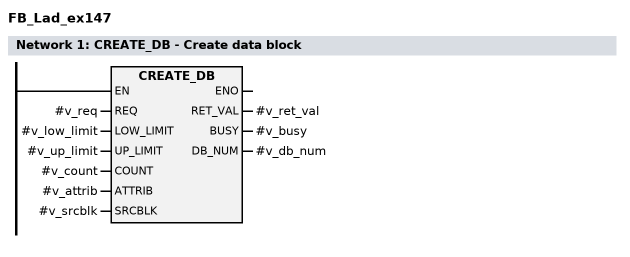
   #v_ret_val := CREATE_DB(REQ := #v_req,
                           LOW_LIMIT := #v_low_limit,
                           UP_LIMIT := #v_up_limit,
                           COUNT := #v_count,
                           ATTRIB := #v_attrib,
                           SRCBLK := #v_srcblk,
                           BUSY => #v_busy,
                           DB_NUM => #v_db_num);
END_REGION
END_FUNCTION_BLOCK

FUNCTION_BLOCK "FB_Lad_ex150"   // FB54, LAD
{ S7_Optimized_Access := 'TRUE' }
   VAR_INPUT
      v_req : Bool;
      v_db_number : DB_ANY;
   END_VAR
   VAR_OUTPUT
      v_ret_val : Int;
      v_db_length : UDInt;
      v_attrib : Byte;
   END_VAR
BEGIN

REGION Network 1: ATTR_DB - Read data block attribute
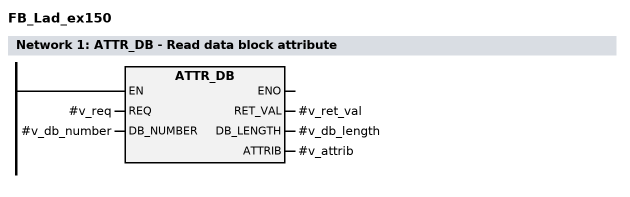
   #v_ret_val := ATTR_DB(REQ := #v_req,
                         DB_NUMBER := #v_db_number,
                         DB_LENGTH => #v_db_length,
                         ATTRIB => #v_attrib);
END_REGION
END_FUNCTION_BLOCK

FUNCTION_BLOCK "FB_Lad_ex151"   // FB55, LAD
{ S7_Optimized_Access := 'TRUE' }
   VAR_INPUT
      v_req : Bool;
      v_db_number : UInt;
   END_VAR
   VAR_OUTPUT
      v_ret_val : Int;
      v_busy : Bool;
   END_VAR
BEGIN

REGION Network 1: DELETE_DB - Delete data block
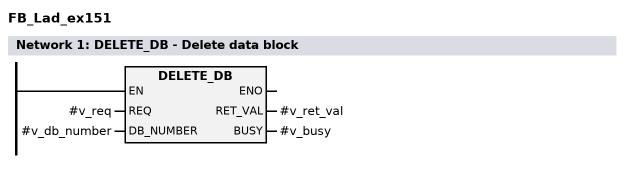
   #v_ret_val := DELETE_DB(REQ := #v_req, DB_NUMBER := #v_db_number, BUSY => #v_busy);
END_REGION
END_FUNCTION_BLOCK

FUNCTION_BLOCK "FB_Lad_ex154"   // FB56, LAD
{ S7_Optimized_Access := 'TRUE' }
   VAR_INPUT
      v_ioid : Byte;
      v_addr : Word;
      v_ret_val : Int;
   END_VAR
   VAR_OUTPUT
      v_hwid : Hw_Io;
   END_VAR
BEGIN

REGION Network 1: LOG2MOD - Determine the hardware identifier from addressing of STEP 7 V5.5 SPx
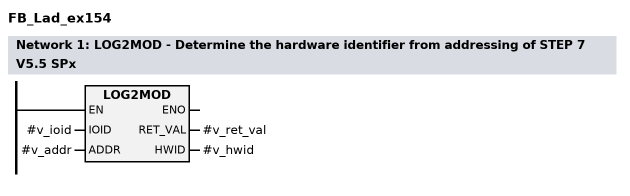
   #v_ret_val := LOG2MOD(IOID := #v_ioid, ADDR := #v_addr, HWID => #v_hwid);
END_REGION
END_FUNCTION_BLOCK

FUNCTION_BLOCK "FB_Lad_ex155"   // FB57, LAD
{ S7_Optimized_Access := 'TRUE' }
   VAR_INPUT
      v_addr : Variant;
      v_ret_val : Int;
   END_VAR
   VAR_OUTPUT
      v_laddr : Hw_Io;
   END_VAR
BEGIN

REGION Network 1: IO2MOD - Determine hardware identifier from an IO address
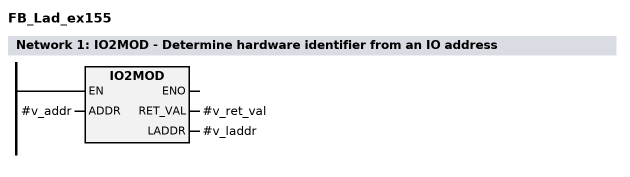
   #v_ret_val := IO2MOD(ADDR := #v_addr, LADDR => #v_laddr);
END_REGION
END_FUNCTION_BLOCK

FUNCTION_BLOCK "FB_Lad_ex156"   // FB58, LAD
{ S7_Optimized_Access := 'TRUE' }
   VAR_INPUT
      v_laddr : Hw_Io;
      v_ret_val : Int;
   END_VAR
   VAR_OUTPUT
      v_piaddr : UDInt;
      v_picount : UInt;
      v_pqaddr : UDInt;
      v_pqcount : UInt;
   END_VAR
BEGIN

REGION Network 1: RD_ADDR - Determine IO addresses from the hardware identifier
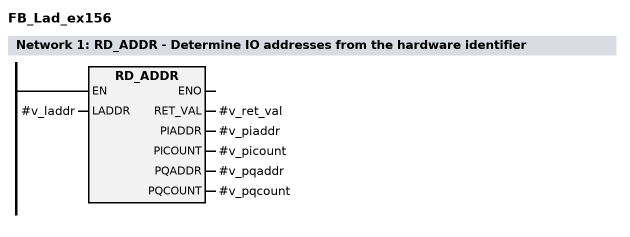
   #v_ret_val := RD_ADDR(LADDR := #v_laddr,
                         PIADDR => #v_piaddr,
                         PICount => #v_picount,
                         PQADDR => #v_pqaddr,
                         PQCount => #v_pqcount);
END_REGION
END_FUNCTION_BLOCK

FUNCTION_BLOCK "FB_Lad_ex157"   // FB59, LAD
{ S7_Optimized_Access := 'TRUE' }
   VAR_INPUT
      v_master : Int;
      v_station : Int;
      v_slot : Int;
      v_subslot : Int;
      v_ret_val : Int;
   END_VAR
   VAR_OUTPUT
      v_laddr : Hw_Io;
   END_VAR
BEGIN

REGION Network 1: GEO_LOG - Determine hardware identifier from slot
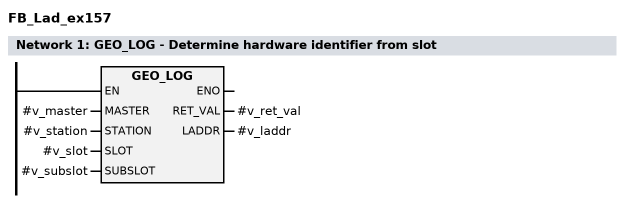
   #v_ret_val := GEO_LOG(MASTER := #v_master,
                         STATION := #v_station,
                         SLOT := #v_slot,
                         SUBSLOT := #v_subslot,
                         LADDR => #v_laddr);
END_REGION
END_FUNCTION_BLOCK

FUNCTION_BLOCK "FB_Lad_ex158"   // FB60, LAD
{ S7_Optimized_Access := 'TRUE' }
   VAR_INPUT
      v_laddr : Hw_Io;
      v_ret_val : Int;
   END_VAR
   VAR_OUTPUT
      v_area : Int;
      v_master : Int;
      v_station : Int;
      v_slot : Int;
      v_subslot : Int;
      v_offset : Int;
   END_VAR
BEGIN

REGION Network 1: LOG_GEO - Determine slot from hardware identifier
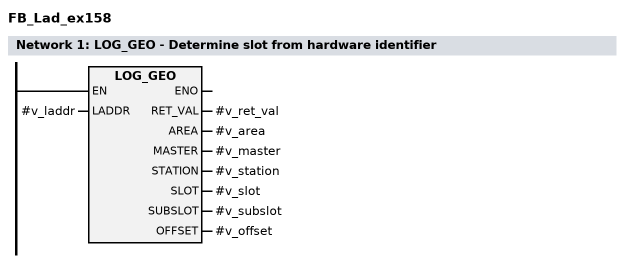
   #v_ret_val := LOG_GEO(LADDR := #v_laddr,
                         AREA => #v_area,
                         MASTER => #v_master,
                         STATION => #v_station,
                         SLOT => #v_slot,
                         SUBSLOT => #v_subslot,
                         OFFSET => #v_offset);
END_REGION
END_FUNCTION_BLOCK

FUNCTION_BLOCK "FB_Lad_ex160"   // FB61, LAD
{ S7_Optimized_Access := 'TRUE' }
   VAR_INPUT
      v_subnetid : Byte;
      v_rack : Word;
      v_slot : Word;
      v_subslot : Byte;
      v_subaddr : Word;
      v_ret_val : Int;
   END_VAR
   VAR_OUTPUT
      v_ioid : Byte;
      v_laddr : Hw_Module;
   END_VAR
BEGIN

REGION Network 1: GADR_LGC - Determine hardware identifier from slot and offset in the user data address area
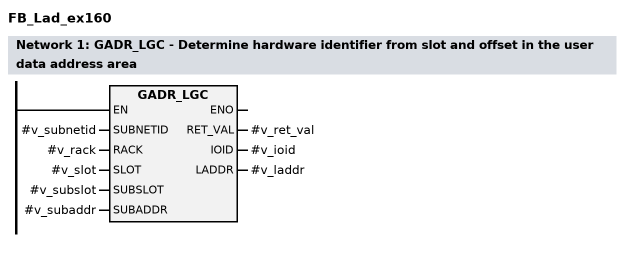
   #v_ret_val := GADR_LGC(SUBNETID := #v_subnetid,
                          RACK := #v_rack,
                          SLOT := #v_slot,
                          SUBSLOT := #v_subslot,
                          SUBADDR := #v_subaddr,
                          IOID => #v_ioid,
                          LADDR => #v_laddr);
END_REGION
END_FUNCTION_BLOCK

FUNCTION_BLOCK "FB_Lad_ex161"   // FB62, LAD
{ S7_Optimized_Access := 'TRUE' }
   VAR_INPUT
      v_ioid : Byte;
      v_laddr : Hw_Module;
      v_ret_val : Int;
   END_VAR
   VAR_OUTPUT
      v_area : Byte;
      v_rack : Word;
      v_slot : Word;
      v_subaddr : Word;
   END_VAR
BEGIN

REGION Network 1: LGC_GADR - Determine slot from hardware identifier
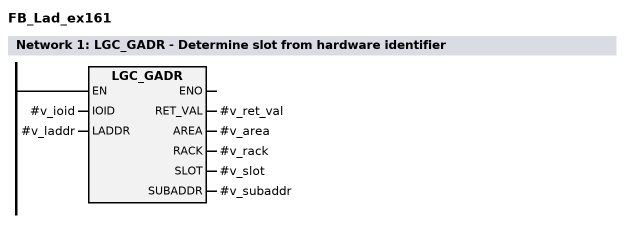
   #v_ret_val := LGC_GADR(IOID := #v_ioid,
                          LADDR := #v_laddr,
                          AREA => #v_area,
                          RACK => #v_rack,
                          SLOT => #v_slot,
                          SUBADDR => #v_subaddr);
END_REGION
END_FUNCTION_BLOCK

FUNCTION_BLOCK "FB_Lad_ws001"   // FB63, LAD
{ S7_Optimized_Access := 'TRUE' }
   VAR_INPUT
      v_ctrl_db : DB_WWW;
   END_VAR
   VAR_OUTPUT
      v_ret_val : Int;
   END_VAR
BEGIN

REGION Network 1: WWW - Synchronizing user pages
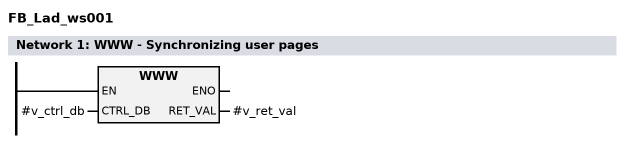
   #v_ret_val := WWW(CTRL_DB := #v_ctrl_db);
END_REGION
END_FUNCTION_BLOCK

FUNCTION_BLOCK "FB_Lad_ex025"   // FB64, LAD
{ S7_Optimized_Access := 'TRUE' }
   VAR_INPUT
      v_n : Int;
      v_ret_val : Word;
   END_VAR
   VAR_IN_OUT
      v_in : Variant;
      v_out : Variant;
   END_VAR
BEGIN

REGION Network 1: ATH - Convert ASCII string to hexadecimal number
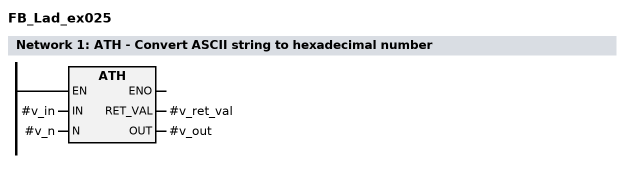
   #v_ret_val := ATH(IN := #v_in, N := #v_n, OUT => #v_out);
END_REGION
END_FUNCTION_BLOCK

FUNCTION_BLOCK "FB_Lad_ex026"   // FB65, LAD
{ S7_Optimized_Access := 'TRUE' }
   VAR_INPUT
      v_n : UInt;
      v_ret_val : Word;
   END_VAR
   VAR_IN_OUT
      v_in : Variant;
      v_out : Variant;
   END_VAR
BEGIN

REGION Network 1: HTA - Convert hexadecimal number to ASCII string
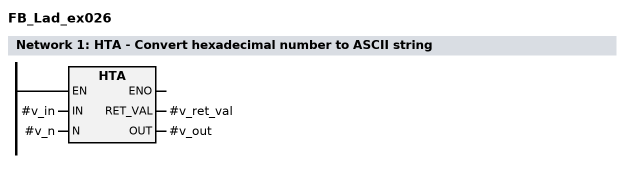
   #v_ret_val := HTA(IN := #v_in, N := #v_n, OUT => #v_out);
END_REGION
END_FUNCTION_BLOCK

FUNCTION_BLOCK "FB_Lad_ex036"   // FB66, LAD
{ S7_Optimized_Access := 'TRUE' }
   VAR_INPUT
      v_size : DInt;
      v_out : WString;
   END_VAR
   VAR_IN_OUT
      v_variable : Array[0..99] of Byte;
   END_VAR
BEGIN

REGION Network 1: GetSymbolName - Read out a tag on the input parameter
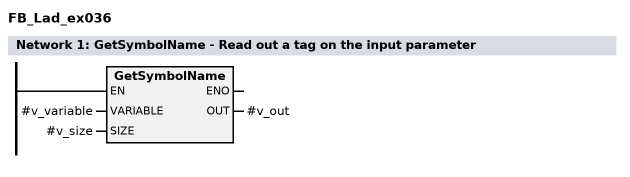
   // no SCL statement known for GetSymbolName: written as a call
   #v_out := GetSymbolName(variable := #v_variable, size := #v_size);
END_REGION
END_FUNCTION_BLOCK

FUNCTION_BLOCK "FB_Lad_ex060"   // FB67, LAD
{ S7_Optimized_Access := 'TRUE' }
   VAR_INPUT
      v_laddr : Hw_Io;
      v_ret_val : Int;
   END_VAR
   VAR_IN_OUT
      v_record : Variant;
   END_VAR
BEGIN

REGION Network 1: DPRD_DAT - Read consistent data of a DP standard slave
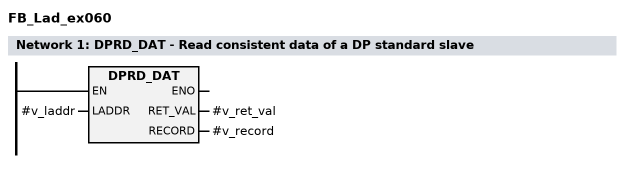
   #v_ret_val := DPRD_DAT(LADDR := #v_laddr, RECORD => #v_record);
END_REGION
END_FUNCTION_BLOCK

FUNCTION_BLOCK "FB_Lad_ex065"   // FB68, LAD
{ S7_Optimized_Access := 'TRUE' }
   VAR_INPUT
      v_req : Bool;
      v_laddr : Hw_DpSlave;
      v_ret_val : DInt;
   END_VAR
   VAR_OUTPUT
      v_busy : Bool;
   END_VAR
   VAR_IN_OUT
      v_record : Variant;
   END_VAR
BEGIN

REGION Network 1: DPNRM_DG - Read diagnostics data from a DP slave
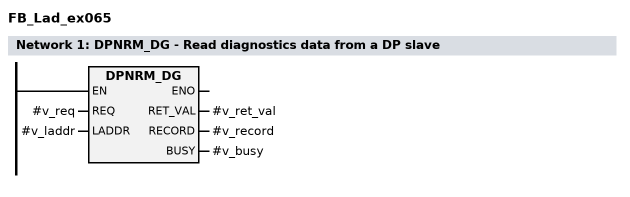
   #v_ret_val := DPNRM_DG(REQ := #v_req, LADDR := #v_laddr, RECORD => #v_record, BUSY => #v_busy);
END_REGION
END_FUNCTION_BLOCK

FUNCTION_BLOCK "FB_Lad_ex097"   // FB69, LAD
{ S7_Optimized_Access := 'TRUE' }
   VAR_INPUT
      v_req : Bool;
      v_laddr : Hw_Io;
      v_recnum : Byte;
      v_ret_val : Int;
   END_VAR
   VAR_OUTPUT
      v_busy : Bool;
   END_VAR
   VAR_IN_OUT
      v_record : Variant;
   END_VAR
BEGIN

REGION Network 1: RD_DPARA - Read module data record asynchronously
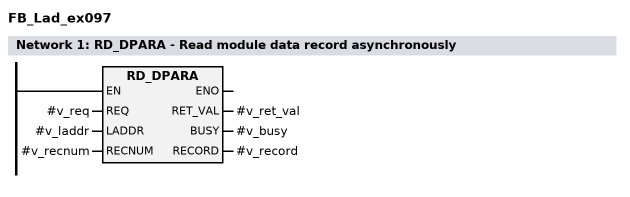
   #v_ret_val := RD_DPARA(REQ := #v_req,
                          LADDR := #v_laddr,
                          RECNUM := #v_recnum,
                          BUSY => #v_busy,
                          RECORD => #v_record);
END_REGION
END_FUNCTION_BLOCK

FUNCTION_BLOCK "FB_Lad_ex098"   // FB70, LAD
{ S7_Optimized_Access := 'TRUE' }
   VAR_INPUT
      v_ioid : Byte;
      v_laddr : Hw_Io;
      v_recnum : Byte;
      v_ret_val : Int;
   END_VAR
   VAR_IN_OUT
      v_record : Variant;
   END_VAR
BEGIN

REGION Network 1: RD_DPARM - Read data record from configured system data
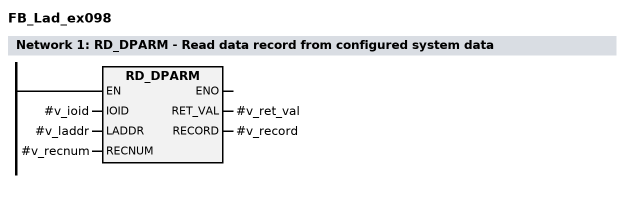
   #v_ret_val := RD_DPARM(IOID := #v_ioid, LADDR := #v_laddr, RECNUM := #v_recnum, RECORD => #v_record);
END_REGION
END_FUNCTION_BLOCK

FUNCTION_BLOCK "FB_Lad_ex124"   // FB71, LAD
{ S7_Optimized_Access := 'TRUE' }
   VAR_INPUT
      v_ret_val : Int;
   END_VAR
   VAR_IN_OUT
      v_top_si : Array[0..99] of Byte;
      v_start_up_si : Array[0..99] of Byte;
   END_VAR
BEGIN

REGION Network 1: RD_SINFO - Read current OB start information
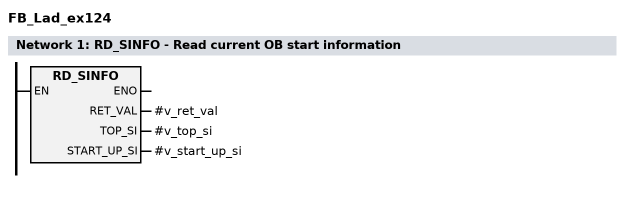
   #v_ret_val := RD_SINFO(TOP_SI => #v_top_si, START_UP_SI => #v_start_up_si);
END_REGION
END_FUNCTION_BLOCK

FUNCTION_BLOCK "FB_Lad_ex148"   // FB72, LAD
{ S7_Optimized_Access := 'TRUE' }
   VAR_INPUT
      v_req : Bool;
      v_ret_val : Int;
   END_VAR
   VAR_OUTPUT
      v_busy : Bool;
   END_VAR
   VAR_IN_OUT
      v_srcblk : Variant;
      v_dstblk : Variant;
   END_VAR
BEGIN

REGION Network 1: READ_DBL - Read from data block in the load memory
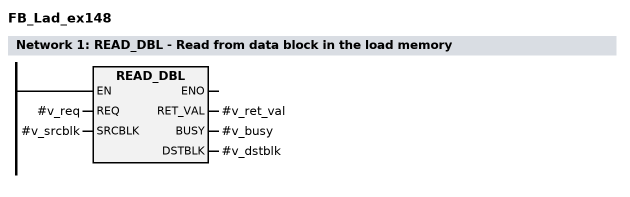
   #v_ret_val := READ_DBL(REQ := #v_req, SRCBLK := #v_srcblk, BUSY => #v_busy, DSTBLK => #v_dstblk);
END_REGION
END_FUNCTION_BLOCK

FUNCTION_BLOCK "FB_Lad_ex149"   // FB73, LAD
{ S7_Optimized_Access := 'TRUE' }
   VAR_INPUT
      v_req : Bool;
      v_ret_val : Int;
   END_VAR
   VAR_OUTPUT
      v_busy : Bool;
   END_VAR
   VAR_IN_OUT
      v_srcblk : Variant;
      v_dstblk : Variant;
   END_VAR
BEGIN

REGION Network 1: WRIT_DBL - Write to data block in the load memory
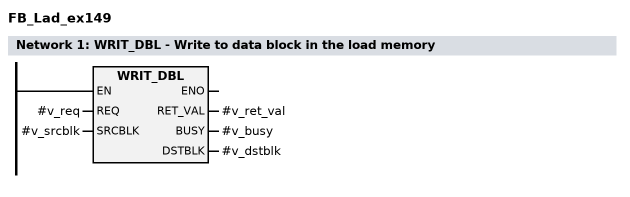
   #v_ret_val := WRIT_DBL(REQ := #v_req, SRCBLK := #v_srcblk, BUSY => #v_busy, DSTBLK => #v_dstblk);
END_REGION
END_FUNCTION_BLOCK

FUNCTION_BLOCK "FB_Lad_ou010"   // FB74, LAD
{ S7_Optimized_Access := 'TRUE' }
   VAR_INPUT
      v_req : Bool;
      v_id : Conn_Ouc;
   END_VAR
   VAR_OUTPUT
      v_done : Bool;
      v_busy : Bool;
      v_error : Bool;
      v_status : Word;
   END_VAR
   VAR_IN_OUT
      v_connect : TCON_Param;
   END_VAR
   VAR
      inst : TCON;
   END_VAR
BEGIN

REGION Network 1: TCON - Establish communication connection
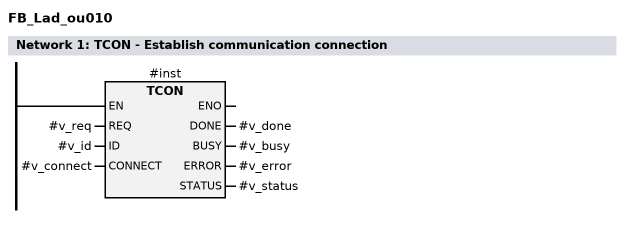
   #inst(REQ := #v_req,   // TCON
         ID := #v_id,
         CONNECT := #v_connect,
         DONE => #v_done,
         BUSY => #v_busy,
         ERROR => #v_error,
         STATUS => #v_status);
END_REGION
END_FUNCTION_BLOCK

FUNCTION_BLOCK "FB_Lad_ou002"   // FB75, LAD
{ S7_Optimized_Access := 'TRUE' }
   VAR_INPUT
      v_req : Bool;
      v_cont : Bool;
      v_len : UDInt;
   END_VAR
   VAR_OUTPUT
      v_done : Bool;
      v_busy : Bool;
      v_error : Bool;
      v_status : Word;
   END_VAR
   VAR_IN_OUT
      v_connect : Array[0..99] of Byte;
      v_data : Array[0..99] of Byte;
      v_addr : Array[0..99] of Byte;
      v_com_rst : Bool;
   END_VAR
   VAR
      inst : TSEND_C;
   END_VAR
BEGIN

REGION Network 1: TSEND_C - Establishing a connection and sending data
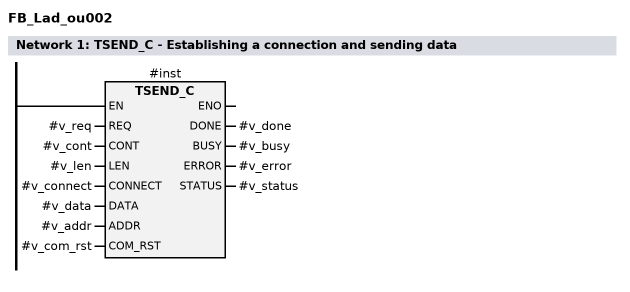
   #inst(REQ := #v_req,   // TSEND_C
         CONT := #v_cont,
         LEN := #v_len,
         CONNECT := #v_connect,
         DATA := #v_data,
         ADDR := #v_addr,
         COM_RST := #v_com_rst,
         DONE => #v_done,
         BUSY => #v_busy,
         ERROR => #v_error,
         STATUS => #v_status);
END_REGION
END_FUNCTION_BLOCK

FUNCTION_BLOCK "FB_Lad_ou004"   // FB76, LAD
{ S7_Optimized_Access := 'TRUE' }
   VAR_INPUT
      v_en_r : Bool;
      v_cont : Bool;
      v_len : UDInt;
      v_adhoc : Bool;
   END_VAR
   VAR_OUTPUT
      v_done : Bool;
      v_busy : Bool;
      v_error : Bool;
      v_status : Word;
      v_rcvd_len : UDInt;
   END_VAR
   VAR_IN_OUT
      v_connect : Array[0..99] of Byte;
      v_data : Array[0..99] of Byte;
      v_addr : Array[0..99] of Byte;
      v_com_rst : Bool;
   END_VAR
   VAR
      inst : TRCV_C;
   END_VAR
BEGIN

REGION Network 1: TRCV_C - Establishing a connection and receiving data
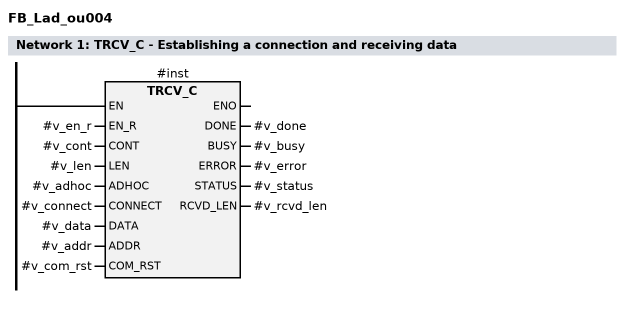
   #inst(EN_R := #v_en_r,   // TRCV_C
         CONT := #v_cont,
         LEN := #v_len,
         ADHOC := #v_adhoc,
         CONNECT := #v_connect,
         DATA := #v_data,
         ADDR := #v_addr,
         COM_RST := #v_com_rst,
         DONE => #v_done,
         BUSY => #v_busy,
         ERROR => #v_error,
         STATUS => #v_status,
         RCVD_LEN => #v_rcvd_len);
END_REGION
END_FUNCTION_BLOCK

FUNCTION_BLOCK "FB_Lad_ou011"   // FB77, LAD
{ S7_Optimized_Access := 'TRUE' }
   VAR_INPUT
      v_req : Bool;
      v_id : Conn_Ouc;
   END_VAR
   VAR_OUTPUT
      v_done : Bool;
      v_busy : Bool;
      v_error : Bool;
      v_status : Word;
   END_VAR
   VAR_IN_OUT
      v_connect : Array[0..99] of Byte;
   END_VAR
   VAR
      inst : TCON;
   END_VAR
BEGIN

REGION Network 1: TCON - Establish communication connection
